// TIA Portal V20 export
VAR_GLOBAL   // PLC tag table "Standard-Variablentabelle"
   System_Byte AT %MB1001 : Byte;
   FirstScan AT %M1001.0 : Bool;
   DiagStatusUpdate AT %M1001.1 : Bool;
   AlwaysTRUE AT %M1001.2 : Bool;
   AlwaysFALSE AT %M1001.3 : Bool;
   Clock_Byte AT %MB1000 : Byte;
   Clock_10Hz AT %M1000.0 : Bool;
   Clock_5Hz AT %M1000.1 : Bool;
   "Clock_2.5Hz" AT %M1000.2 : Bool;
   Clock_2Hz AT %M1000.3 : Bool;
   "Clock_1.25Hz" AT %M1000.4 : Bool;
   Clock_1Hz AT %M1000.5 : Bool;
   "Clock_0.625Hz" AT %M1000.6 : Bool;
   "Clock_0.5Hz" AT %M1000.7 : Bool;
   IBS0 AT %M0.2 : Bool;   // Immer 0, muss nach Inbetriebnahme entfernt werden !!!
   IBS1 AT %M0.3 : Bool;   // immer1, muss nach Inbetriebnahme entfernt werden !!!
   "Zyklisch wechselnder Merker" AT %M70.6 : Bool;
   DA_Anlagenzustand_Trigger_2 AT %Q0.1 : Bool;   // DA +SK2-481P1 Signalbeleuchtung Trigger 2
   DA_0_3 AT %Q0.3 : Bool;
   DA_Anlagenbeleuchtung AT %Q0.4 : Bool;   // DA +SK2-481P1 Signalbeleuchtung Trigger 3 LED Weiß
   "DA_Selektivmodul Reset" AT %Q0.6 : Bool;   // DA +SK2-323T1 Selektivmodul 24V Reset
   DA_0_7 AT %Q0.7 : Bool;
   DA_0_2 AT %Q0.2 : Bool;
   DA_Anlagenzustand_Trigger_1 AT %Q0.0 : Bool;   // DA +SK2-481P1 Signalbeleuchtung Trigger 1
   DA_0_5 AT %Q0.5 : Bool;
   "Ablauf aktiv" AT %M1.7 : Bool;
   Simulation_DE200_bis_DE2199 AT %I200.0 : "DataRange";   // Simulation DE200 bis DE2199
   FL_Clock_1Hz AT %M1004.0 : Bool;
   HM_Clock_1Hz AT %M1004.1 : Bool;
   "DA_Bedienerkonsole_Front_LED_K0-K7_ROT" AT %QB20 : Byte;   // +SK2-458K2 Bedienerkonsole LED K0 - K7 Farbe ROT
   "DA_Bedienerkonsole_Front_LED_K0-K7_GRÜN" AT %QB21 : Byte;   // +SK2-458K2 Bedienerkonsole LED K0 - K7 Farbe GRÜN
   "DA_Bedienerkonsole_Front_LED_K0-K7_BLAU" AT %QB22 : Byte;   // +SK2-458K2 Bedienerkonsole LED K0 - K7 Farbe BLAU
   "NOP" AT %M0.4 : Bool;   // NOP, Dummy keine Funktion
   DA_Extern_OUT1 AT %Q1.0 : Bool;   // DA +SK2-483PK1 Externe Schnittstelle an Messgerät
   DA_Extern_OUT2 AT %Q1.1 : Bool;   // DA +SK2-483PK2 Externe Schnittstelle an Messgerät
   DA_Extern_OUT3 AT %Q1.2 : Bool;   // DA +SK2-483PK3 Externe Schnittstelle an Messgerät
   DA_Extern_OUT4 AT %Q1.3 : Bool;   // DA +SK2-483PK4 Externe Schnittstelle an Messgerät
   DA_1_4 AT %Q1.4 : Bool;
   DA_1_5 AT %Q1.5 : Bool;
   DA_1_6 AT %Q1.6 : Bool;
   DA_1_7 AT %Q1.7 : Bool;
   TEST AT %M500.4 : Bool;
   Tag_1 AT %I206.0 : Bool;
   Tag_2 AT %M5000.1 : Bool;
END_VAR
